TYPE ST_AlarmOut :
STRUCT
	arbFatalError			:ARRAY[0..nALARM_MAX_NO] OF ST_AlarmProperties;
	arbError				:ARRAY[0..nALARM_MAX_NO] OF ST_AlarmProperties;
	arbWarning			:ARRAY[0..nALARM_MAX_NO] OF ST_AlarmProperties;
	arbMessage			:ARRAY[0..nALARM_MAX_NO] OF ST_AlarmProperties;
	arbHint				:ARRAY[0..nALARM_MAX_NO] OF ST_AlarmProperties;
	bFatalError			:BOOL;				(* Fatal error in group / Fataler Fehler in der Gruppe *)
	bError				:BOOL;				(* Error in group / Fehler in der Gruppe *)
	bWarning			:BOOL;				(* Warning in group / Warnung  in der Gruppe *)
	bMessage			:BOOL;				(* Message in group / Meldung in der Gruppe *)
	bHint				:BOOL;				(* Hint in group / Hint in der Gruppe *)
END_STRUCT
END_TYPE

(* stored: Version 1.1.0.1, ProductVersion 3.1.4024.15
   DUT ST_AlarmOut: Id {f2fabadd-deca-4973-a49f-56d31c58f4bb} *)
